// TIA Portal V20 export
// export: Created 2026-10-20T12:44:59.1372721Z, ExportSetting WithDefaults, DisplayName Totally Integrated Automation Portal, DisplayVersion V20 Update 6, DisplayName TIA Portal Openness, DisplayVersion V20 Update 6, DisplayName TIA Portal Version Control Interface, DisplayVersion V20 Update 6, DisplayName SINAMICS Startdrive Advanced, DisplayVersion V20 SP1, DisplayName SINAMICS Startdrive G130, G150, S120, S150, SINAMICS MV, G220, S200, S210, DisplayVersion V20 SP1, DisplayName SINAMICS Startdrive G110M, G120, G120C, G120D, G120P, G115D, DisplayVersion V20 SP1, DisplayName STEP 7 Professional, DisplayVersion V20 Update 6, DisplayName STEP 7 Safety, DisplayVersion V20 Update 2, DisplayName WinCC Basic/Comfort/Advanced, DisplayVersion V20 Update 6, DisplayName WinCC Unified, DisplayVersion V20 Update 6
FUNCTION "CNV_Charge_Settings_FC_1" : Void   // FC59, SCL
{ S7_Optimized_Access := 'TRUE' }
VERSION : 0.1
// stored: AutoNumber true, IsIECCheckEnabled false, SetENOAutomatically false, UDAEnableTagReadback false
   VAR_INPUT
      Sys_No : UInt;
      HMI_Box : UInt;
   END_VAR
   VAR_TEMP
      Level : UInt;
   END_VAR
BEGIN
   #Level := #HMI_Box MOD 10;
   "PopUps_DB_1"."ECnv_Settings"[#Sys_No] := "Settings_DB".ECnv_Sys[#Sys_No];

   CASE #Level OF
       1:
           "PopUps_DB_1"."Buffer_Cnv_Settings_1"[#Sys_No] := "Settings_DB".LCnv_Sys[#Sys_No].Cnv_Level[1].Cnv1;
           "PopUps_DB_1"."Buffer_Cnv_Settings_2"[#Sys_No] := "Settings_DB".LCnv_Sys[#Sys_No].Cnv_Level[1].Cnv2;
       2:
           "PopUps_DB_1"."Buffer_Cnv_Settings_1"[#Sys_No] := "Settings_DB".LCnv_Sys[#Sys_No].Cnv_Level[2].Cnv1;
           "PopUps_DB_1"."Buffer_Cnv_Settings_2"[#Sys_No] := "Settings_DB".LCnv_Sys[#Sys_No].Cnv_Level[2].Cnv2;
       3:
           "PopUps_DB_1"."Buffer_Cnv_Settings_1"[#Sys_No] := "Settings_DB".LCnv_Sys[#Sys_No].Cnv_Level[3].Cnv1;
           "PopUps_DB_1"."Buffer_Cnv_Settings_2"[#Sys_No] := "Settings_DB".LCnv_Sys[#Sys_No].Cnv_Level[3].Cnv2;
       4:
           "PopUps_DB_1"."Buffer_Cnv_Settings_1"[#Sys_No] := "Settings_DB".LCnv_Sys[#Sys_No].Cnv_Level[4].Cnv1;
           "PopUps_DB_1"."Buffer_Cnv_Settings_2"[#Sys_No] := "Settings_DB".LCnv_Sys[#Sys_No].Cnv_Level[4].Cnv2;
       5:
           "PopUps_DB_1"."Buffer_Cnv_Settings_1"[#Sys_No] := "Settings_DB".LCnv_Sys[#Sys_No].Cnv_Level[5].Cnv1;
           "PopUps_DB_1"."Buffer_Cnv_Settings_2"[#Sys_No] := "Settings_DB".LCnv_Sys[#Sys_No].Cnv_Level[5].Cnv2;
       6:
           "PopUps_DB_1"."Buffer_Cnv_Settings_1"[#Sys_No] := "Settings_DB".LCnv_Sys[#Sys_No].Cnv_Level[6].Cnv1;
           "PopUps_DB_1"."Buffer_Cnv_Settings_2"[#Sys_No] := "Settings_DB".LCnv_Sys[#Sys_No].Cnv_Level[6].Cnv2;
       7:
           "PopUps_DB_1"."Buffer_Cnv_Settings_1"[#Sys_No] := "Settings_DB".LCnv_Sys[#Sys_No].Cnv_Level[7].Cnv1;
           "PopUps_DB_1"."Buffer_Cnv_Settings_2"[#Sys_No] := "Settings_DB".LCnv_Sys[#Sys_No].Cnv_Level[7].Cnv2;
       8:
           "PopUps_DB_1"."Buffer_Cnv_Settings_1"[#Sys_No] := "Settings_DB".LCnv_Sys[#Sys_No].Cnv_Level[8].Cnv1;
           "PopUps_DB_1"."Buffer_Cnv_Settings_2"[#Sys_No] := "Settings_DB".LCnv_Sys[#Sys_No].Cnv_Level[8].Cnv2;
   END_CASE;
END_FUNCTION
